(*
SPDX-FileCopyrightText: c 2026 Oleksandr Tiutyk <trofimich@gmail.com>
SPDX-License-Identifier: MIT
License: https://opensource.org/license/mit
*)

(*!
<summary>Groups byte-string formatting, editing, search and splitter contracts.</summary>
<description>
Owns the independent child instances and their fixed registration array. Use from one PLC task at a stable address.
</description>
*)

{attribute 'no_assign'}
{attribute 'no_explicit_call' := 'do not call this function block directly'}
FUNCTION_BLOCK StringsTestGroup EXTENDS TOF_Testing.TestGroup<10>
VAR_STAT
	{attribute 'hide'}
	_ClassName : STRING := __POUNAME();
END_VAR
VAR
	_AnyToStringFit255 : StringFitFormattingTest(name := "AnyToStringFit255", parent := THIS^);
	_Append : StringAppendTest(name := "Append", parent := THIS^);
	_AppendFit : StringAppendFitTest(name := "AppendFit", parent := THIS^);
	_ConcatFit255 : StringConcatFitTest(name := "ConcatFit255", parent := THIS^);
	_Contains : StringContainsTest(name := "Contains", parent := THIS^);
	_Join : StringJoinTest(name := "Join", parent := THIS^);
	_ReplaceInSource : StringReplacementTest(name := "ReplaceInSource", parent := THIS^);
	_Split : StringSplitTest(name := "Split", parent := THIS^);
	_Trim : StringTrimTest(name := "Trim", parent := THIS^);
	_SplitterSeparatorBounds : StringSeparatorBoundsTest(name := "SplitterSeparatorBounds", parent := THIS^);

	_Children : ARRAY [0.._ChildCount - 1] OF TOF_Testing.ITestElement :=
	[
		_AnyToStringFit255,
		_Append,
		_AppendFit,
		_ConcatFit255,
		_Contains,
		_Join,
		_ReplaceInSource,
		_Split,
		_Trim,
		_SplitterSeparatorBounds
	];
END_VAR

//! <summary>Borrows the fixed child array. Callers must not modify it.</summary>
{attribute 'monitoring' := 'call'}
PROPERTY Children : REFERENCE TO ARRAY [0.._ChildCount - 1] OF TOF_Testing.ITestElement
GET
Children REF= _Children;
END_GET
END_PROPERTY

//! <summary>Borrows the concrete class name. Callers must not modify it.</summary>
{attribute 'monitoring' := 'call'}
PROPERTY ClassName : REFERENCE TO STRING
GET
ClassName REF= _ClassName;
END_GET
END_PROPERTY

//! <summary>Borrows the compiler-initialized namespace name. Callers must not modify it.</summary>
{attribute 'monitoring' := 'call'}
PROPERTY NamespaceName : REFERENCE TO STRING
GET
NamespaceName REF= CurrentNamespace.Name;
END_GET
END_PROPERTY

//! <summary>Reports the concrete instance size in bytes.</summary>
{attribute 'monitoring' := 'call'}
PROPERTY SelfSize : ULINT
GET
SelfSize := XSIZEOF(THIS^);
END_GET
END_PROPERTY

END_FUNCTION_BLOCK

(* stored: Version 1.1.0.1
   POU StringsTestGroup: Id {19b3bce0-2b8a-49f6-8577-68a0ce66d979}, SpecialFunc None
   Property Children: Id {3920885b-cf79-429d-8649-95fcd197d5e1}
   Get Get: Id {e2f52323-7683-4397-b906-76656b6fb43d}
   Property ClassName: Id {b0cbaaeb-9e33-4526-8daf-61d9aacc9001}
   Get Get: Id {9456c479-a33d-4d23-9b0d-83d72fab0105}
   Property NamespaceName: Id {ee72c81b-6f6b-4481-840e-ff60701d55f7}
   Get Get: Id {05fef4ed-457f-4fa7-837e-f2fd158d4075}
   Property SelfSize: Id {3ef79b4e-f1b5-4120-8334-27aa18f33d76}
   Get Get: Id {726bc39c-6334-4bf4-984d-044a7afaa249} *)
